(*
SPDX-FileCopyrightText: © 2026 Oleksandr Tiutyk <trofimich@gmail.com>
SPDX-License-Identifier: MIT
License: https://opensource.org/license/mit
*)

(*!
<summary>Provides fluent assertions on a copied TIME_OF_DAY value.</summary>
<description>
Copies actual into persistent instance storage before the entry method returns; literals and expression
results therefore remain valid throughout the immediate chain. Owns no heap allocation or pointed-to resource.
The message prefixes every failure until the next preparation. Finish one chain before starting another on
the owning Assertions provider. Use only from the owning test callback on one task, without reentry.
Obtain this context from the owning provider; direct unprepared use is unsupported.
Expected arguments use the declared IEC type; ordinary compiler conversions happen before comparison.
This context does not depend on another assertion context.
Object metadata is available before preparation; inherited equality compares instance identity.
Ordering uses the native IEC comparison of time since midnight, without a duration conversion or wrap-around.
</description>
*)

{attribute 'no_explicit_call' := 'do not call this function block directly'}
FUNCTION_BLOCK TimeOfDayAssertionContext EXTENDS TOF_Core.Object
VAR_STAT
	{attribute 'hide'}
	_ClassName : STRING := __POUNAME();
END_VAR
VAR
	_Actual : TIME_OF_DAY;
	_TestCase : ITestCase;
	_Message : WSTRING(255);
END_VAR

(*!
<summary>Provides the implementation class name.</summary>
<description>
Borrowed read-only reference to compiler-initialized storage, valid throughout the instance lifetime.
Do not modify the returned reference; no ownership is transferred.
</description>
*)
{attribute 'monitoring' := 'call'}
PROPERTY ClassName : REFERENCE TO STRING
GET
ClassName REF= _ClassName;
END_GET
END_PROPERTY

(*!
<summary>Asserts that the actual value is strictly greater than expected.</summary>
<description>
Records failure without interrupting the callback; preserves the message for the rest of the chain.
</description>
<param name="expected">Expected value converted by the compiler to TIME_OF_DAY.</param>
*)
METHOD FINAL IsGreaterThan : REFERENCE TO TimeOfDayAssertionContext
VAR_INPUT
	expected : TIME_OF_DAY;
END_VAR
IF _Actual <= expected THEN
	failComparison(
		expected := expected,
		expectation := "Expected value > "
	);
END_IF

IsGreaterThan REF= THIS^;
END_METHOD

(*!
<summary>Asserts that the actual value meets the inclusive lower boundary.</summary>
<description>
Records failure without interrupting the callback; preserves the message for the rest of the chain.
</description>
<param name="expected">Expected value converted by the compiler to TIME_OF_DAY.</param>
*)
METHOD FINAL IsGreaterThanOrEquals : REFERENCE TO TimeOfDayAssertionContext
VAR_INPUT
	expected : TIME_OF_DAY;
END_VAR
IF _Actual < expected THEN
	failComparison(
		expected := expected,
		expectation := "Expected value >= "
	);
END_IF

IsGreaterThanOrEquals REF= THIS^;
END_METHOD

(*!
<summary>Asserts that the actual value is strictly less than expected.</summary>
<description>
Records failure without interrupting the callback; preserves the message for the rest of the chain.
</description>
<param name="expected">Expected value converted by the compiler to TIME_OF_DAY.</param>
*)
METHOD FINAL IsLessThan : REFERENCE TO TimeOfDayAssertionContext
VAR_INPUT
	expected : TIME_OF_DAY;
END_VAR
IF _Actual >= expected THEN
	failComparison(
		expected := expected,
		expectation := "Expected value < "
	);
END_IF

IsLessThan REF= THIS^;
END_METHOD

(*!
<summary>Asserts that the actual value meets the inclusive upper boundary.</summary>
<description>
Records failure without interrupting the callback; preserves the message for the rest of the chain.
</description>
<param name="expected">Expected value converted by the compiler to TIME_OF_DAY.</param>
*)
METHOD FINAL IsLessThanOrEquals : REFERENCE TO TimeOfDayAssertionContext
VAR_INPUT
	expected : TIME_OF_DAY;
END_VAR
IF _Actual > expected THEN
	failComparison(
		expected := expected,
		expectation := "Expected value <= "
	);
END_IF

IsLessThanOrEquals REF= THIS^;
END_METHOD

(*!
<summary>Provides the library namespace.</summary>
<description>
Borrowed read-only reference to the compiler-initialized namespace, valid throughout the instance lifetime.
Do not modify the returned reference; no ownership is transferred.
</description>
*)
{attribute 'monitoring' := 'call'}
PROPERTY NamespaceName : REFERENCE TO STRING
GET
NamespaceName REF= CurrentNamespace.Name;
END_GET
END_PROPERTY

(*!
<summary>Asserts inequality with the expected value.</summary>
<description>
Records failure without interrupting the callback; preserves the message for the rest of the chain.
</description>
<param name="expected">Expected value converted by the compiler to TIME_OF_DAY.</param>
*)
METHOD FINAL NotToBe : REFERENCE TO TimeOfDayAssertionContext
VAR_INPUT
	expected : TIME_OF_DAY;
END_VAR
IF _Actual = expected THEN
	failComparison(
		expected := expected,
		expectation := "Expected value not to be: "
	);
END_IF

NotToBe REF= THIS^;
END_METHOD

(*!
<summary>Copies the actual operand and replaces the chain-wide message.</summary>
<description>
Called by the owning Assertions provider after it verifies the running test case.
No pointer to this method's input storage is retained. The receiver is borrowed until the next preparation;
the owning provider keeps it alive throughout the immediate chain.
</description>
<param name="actual">Value copied into this context.</param>
<param name="testCase">Borrowed failure receiver for the immediate chain.</param>
<param name="message">Copied diagnostic prefix, including empty to clear the previous prefix.</param>
*)
METHOD INTERNAL FINAL Prepare
VAR_INPUT
	actual : TIME_OF_DAY;
	testCase : ITestCase;
	message : WSTRING(255);
END_VAR
_Actual := actual;
_TestCase := testCase;
_Message := message;
END_METHOD

(*!
<summary>Reports the byte size of this concrete instance.</summary>
<description>
Includes inline fields and nested instances, but excludes separately allocated payloads.
Obtaining the size does not transfer ownership or validate an arbitrary address.
</description>
*)
{attribute 'monitoring' := 'call'}
PROPERTY SelfSize : ULINT
GET
SelfSize := XSIZEOF(THIS^);
END_GET
END_PROPERTY

(*!
<summary>Asserts equality with the expected value.</summary>
<description>
Records failure without interrupting the callback; preserves the message for the rest of the chain.
</description>
<param name="expected">Expected value converted by the compiler to TIME_OF_DAY.</param>
*)
METHOD FINAL ToBe : REFERENCE TO TimeOfDayAssertionContext
VAR_INPUT
	expected : TIME_OF_DAY;
END_VAR
IF _Actual <> expected THEN
	failComparison(
		expected := expected,
		expectation := "Expected: "
	);
END_IF

ToBe REF= THIS^;
END_METHOD

(*!
<summary>Formats a failed typed predicate and reports it with the chain message.</summary>
<description>
Does not change operands or chain state. The receiver retains its first failure. Reporting exceptions
propagate to the enclosing test callback handler; an unprepared receiver is a configuration error.
</description>
<param name="expected">Typed expected operand used only for this diagnostic.</param>
<param name="expectation">Prefix identifying the failed predicate.</param>
*)
METHOD PRIVATE failComparison
VAR_INPUT
	expected : TIME_OF_DAY;
	expectation : WSTRING(40);
END_VAR
VAR
	actualText : WSTRING(255);
	expectedText : WSTRING(255);
	diagnostic : TOF_Core.ERROR_MESSAGE;
END_VAR
actualText := TO_WSTRING(_Actual);
expectedText := TO_WSTRING(expected);

diagnostic := TOF_Core.WideStrings.Concat255(
	expectation,
	expectedText,
	", but was: ",
	actualText
);

TestServices.ReportAssertionFailure(
	testCase := _TestCase,
	message := _Message,
	sourceClassName := ClassName,
	defaultMessage := diagnostic
);
END_METHOD

END_FUNCTION_BLOCK

(* stored: Version 1.1.0.1
   POU TimeOfDayAssertionContext: Id {c2f32a17-d6bb-4e77-a0c7-a69764687539}, SpecialFunc None
   Folder Service methods: Id {188c89e9-9da2-41b3-bf24-83912f7b7527}
   Property ClassName: Id {8b309fa6-c0ea-4800-be65-88b7f0747b4a}
   Get Get: Id {49c939af-92ec-4d7f-99be-f8a6d454a73b}
   Method IsGreaterThan: Id {5b20e12d-0dc4-42b2-8054-6f7788cd3c3d}
   Method IsGreaterThanOrEquals: Id {08246edb-71c3-4585-8e4e-2328624e4d54}
   Method IsLessThan: Id {e597b30e-a1f7-43c1-a1c0-4de9a8736c98}
   Method IsLessThanOrEquals: Id {e55ff887-60a2-462d-a642-555600d3bb52}
   Property NamespaceName: Id {3e1b427e-c85b-40d0-bd65-b68724e4df20}
   Get Get: Id {59f962de-a96e-4044-ab9b-d05d5037b670}
   Method NotToBe: Id {49af30df-e992-463a-9cf2-52b08ad8d548}
   Method Prepare: Id {f63b3656-dcaa-4831-9524-832676be2478}
   Property SelfSize: Id {889dd761-67d8-4ab6-aa62-8998009585b5}
   Get Get: Id {db47c14c-a375-484f-b18a-15b74c1a4ba6}
   Method ToBe: Id {6fc31edc-af9a-4d31-9bcc-eddb7fd8237b}
   Method failComparison: Id {633d0426-b6f8-4d5f-a9dc-11aaaa3bd2ed} *)
